(* IEC 61131-3 sources: STAR-PLC-Agent/results/raw/codex_matrix_resume_20261114/codex_deepseek/SELF007/functional/attempt_0001, 1 file *)

(* ---- test_program.st ---- *)
PROGRAM PLC_PRG
VAR
 BenchStep : UDINT := 0;
 BenchCalls : UDINT := 0;
 BenchDone : BOOL := FALSE;
 BenchUut0 : FB_Task;
 BenchUut1 : FB_Task;
 BenchUut2 : FB_Task;
 BenchUut3 : FB_Task;
 BenchUut4 : FB_Task;
 BenchUut5 : FB_Task;
 BenchUut6 : FB_Task;
 BenchUut7 : FB_Task;
 BenchUut8 : FB_Task;
 TraceIn_Demand : ARRAY[0..59] OF BOOL;
 TraceIn_FaultA : ARRAY[0..59] OF BOOL;
 TraceIn_FaultB : ARRAY[0..59] OF BOOL;
 TraceOut_PumpA : ARRAY[0..59] OF BOOL;
 TraceOut_PumpB : ARRAY[0..59] OF BOOL;
 TraceOut_LeadA : ARRAY[0..59] OF BOOL;
END_VAR

IF NOT BenchDone THEN
 CASE BenchStep OF
 0:
   BenchUut0.Demand := FALSE;
   BenchUut0.FaultA := FALSE;
   BenchUut0.FaultB := FALSE;
   TraceIn_Demand[0] := BenchUut0.Demand;
   TraceIn_FaultA[0] := BenchUut0.FaultA;
   TraceIn_FaultB[0] := BenchUut0.FaultB;
   BenchUut0();
   TraceOut_PumpA[0] := BenchUut0.PumpA;
   TraceOut_PumpB[0] := BenchUut0.PumpB;
   TraceOut_LeadA[0] := BenchUut0.LeadA;
   BenchCalls := BenchCalls + 1;
 1:
   BenchUut0.Demand := TRUE;
   BenchUut0.FaultA := FALSE;
   BenchUut0.FaultB := FALSE;
   TraceIn_Demand[1] := BenchUut0.Demand;
   TraceIn_FaultA[1] := BenchUut0.FaultA;
   TraceIn_FaultB[1] := BenchUut0.FaultB;
   BenchUut0();
   TraceOut_PumpA[1] := BenchUut0.PumpA;
   TraceOut_PumpB[1] := BenchUut0.PumpB;
   TraceOut_LeadA[1] := BenchUut0.LeadA;
   BenchCalls := BenchCalls + 1;
 2:
   BenchUut0.Demand := TRUE;
   BenchUut0.FaultA := FALSE;
   BenchUut0.FaultB := FALSE;
   TraceIn_Demand[2] := BenchUut0.Demand;
   TraceIn_FaultA[2] := BenchUut0.FaultA;
   TraceIn_FaultB[2] := BenchUut0.FaultB;
   BenchUut0();
   TraceOut_PumpA[2] := BenchUut0.PumpA;
   TraceOut_PumpB[2] := BenchUut0.PumpB;
   TraceOut_LeadA[2] := BenchUut0.LeadA;
   BenchCalls := BenchCalls + 1;
 3:
   BenchUut0.Demand := FALSE;
   BenchUut0.FaultA := FALSE;
   BenchUut0.FaultB := FALSE;
   TraceIn_Demand[3] := BenchUut0.Demand;
   TraceIn_FaultA[3] := BenchUut0.FaultA;
   TraceIn_FaultB[3] := BenchUut0.FaultB;
   BenchUut0();
   TraceOut_PumpA[3] := BenchUut0.PumpA;
   TraceOut_PumpB[3] := BenchUut0.PumpB;
   TraceOut_LeadA[3] := BenchUut0.LeadA;
   BenchCalls := BenchCalls + 1;
 4:
   BenchUut0.Demand := FALSE;
   BenchUut0.FaultA := FALSE;
   BenchUut0.FaultB := FALSE;
   TraceIn_Demand[4] := BenchUut0.Demand;
   TraceIn_FaultA[4] := BenchUut0.FaultA;
   TraceIn_FaultB[4] := BenchUut0.FaultB;
   BenchUut0();
   TraceOut_PumpA[4] := BenchUut0.PumpA;
   TraceOut_PumpB[4] := BenchUut0.PumpB;
   TraceOut_LeadA[4] := BenchUut0.LeadA;
   BenchCalls := BenchCalls + 1;
 5:
   BenchUut0.Demand := TRUE;
   BenchUut0.FaultA := FALSE;
   BenchUut0.FaultB := FALSE;
   TraceIn_Demand[5] := BenchUut0.Demand;
   TraceIn_FaultA[5] := BenchUut0.FaultA;
   TraceIn_FaultB[5] := BenchUut0.FaultB;
   BenchUut0();
   TraceOut_PumpA[5] := BenchUut0.PumpA;
   TraceOut_PumpB[5] := BenchUut0.PumpB;
   TraceOut_LeadA[5] := BenchUut0.LeadA;
   BenchCalls := BenchCalls + 1;
 6:
   BenchUut0.Demand := FALSE;
   BenchUut0.FaultA := FALSE;
   BenchUut0.FaultB := FALSE;
   TraceIn_Demand[6] := BenchUut0.Demand;
   TraceIn_FaultA[6] := BenchUut0.FaultA;
   TraceIn_FaultB[6] := BenchUut0.FaultB;
   BenchUut0();
   TraceOut_PumpA[6] := BenchUut0.PumpA;
   TraceOut_PumpB[6] := BenchUut0.PumpB;
   TraceOut_LeadA[6] := BenchUut0.LeadA;
   BenchCalls := BenchCalls + 1;
 7:
   BenchUut1.Demand := TRUE;
   BenchUut1.FaultA := TRUE;
   BenchUut1.FaultB := TRUE;
   TraceIn_Demand[7] := BenchUut1.Demand;
   TraceIn_FaultA[7] := BenchUut1.FaultA;
   TraceIn_FaultB[7] := BenchUut1.FaultB;
   BenchUut1();
   TraceOut_PumpA[7] := BenchUut1.PumpA;
   TraceOut_PumpB[7] := BenchUut1.PumpB;
   TraceOut_LeadA[7] := BenchUut1.LeadA;
   BenchCalls := BenchCalls + 1;
 8:
   BenchUut1.Demand := FALSE;
   BenchUut1.FaultA := TRUE;
   BenchUut1.FaultB := TRUE;
   TraceIn_Demand[8] := BenchUut1.Demand;
   TraceIn_FaultA[8] := BenchUut1.FaultA;
   TraceIn_FaultB[8] := BenchUut1.FaultB;
   BenchUut1();
   TraceOut_PumpA[8] := BenchUut1.PumpA;
   TraceOut_PumpB[8] := BenchUut1.PumpB;
   TraceOut_LeadA[8] := BenchUut1.LeadA;
   BenchCalls := BenchCalls + 1;
 9:
   BenchUut1.Demand := TRUE;
   BenchUut1.FaultA := TRUE;
   BenchUut1.FaultB := FALSE;
   TraceIn_Demand[9] := BenchUut1.Demand;
   TraceIn_FaultA[9] := BenchUut1.FaultA;
   TraceIn_FaultB[9] := BenchUut1.FaultB;
   BenchUut1();
   TraceOut_PumpA[9] := BenchUut1.PumpA;
   TraceOut_PumpB[9] := BenchUut1.PumpB;
   TraceOut_LeadA[9] := BenchUut1.LeadA;
   BenchCalls := BenchCalls + 1;
 10:
   BenchUut1.Demand := TRUE;
   BenchUut1.FaultA := FALSE;
   BenchUut1.FaultB := FALSE;
   TraceIn_Demand[10] := BenchUut1.Demand;
   TraceIn_FaultA[10] := BenchUut1.FaultA;
   TraceIn_FaultB[10] := BenchUut1.FaultB;
   BenchUut1();
   TraceOut_PumpA[10] := BenchUut1.PumpA;
   TraceOut_PumpB[10] := BenchUut1.PumpB;
   TraceOut_LeadA[10] := BenchUut1.LeadA;
   BenchCalls := BenchCalls + 1;
 11:
   BenchUut1.Demand := FALSE;
   BenchUut1.FaultA := TRUE;
   BenchUut1.FaultB := TRUE;
   TraceIn_Demand[11] := BenchUut1.Demand;
   TraceIn_FaultA[11] := BenchUut1.FaultA;
   TraceIn_FaultB[11] := BenchUut1.FaultB;
   BenchUut1();
   TraceOut_PumpA[11] := BenchUut1.PumpA;
   TraceOut_PumpB[11] := BenchUut1.PumpB;
   TraceOut_LeadA[11] := BenchUut1.LeadA;
   BenchCalls := BenchCalls + 1;
 12:
   BenchUut2.Demand := TRUE;
   BenchUut2.FaultA := TRUE;
   BenchUut2.FaultB := FALSE;
   TraceIn_Demand[12] := BenchUut2.Demand;
   TraceIn_FaultA[12] := BenchUut2.FaultA;
   TraceIn_FaultB[12] := BenchUut2.FaultB;
   BenchUut2();
   TraceOut_PumpA[12] := BenchUut2.PumpA;
   TraceOut_PumpB[12] := BenchUut2.PumpB;
   TraceOut_LeadA[12] := BenchUut2.LeadA;
   BenchCalls := BenchCalls + 1;
 13:
   BenchUut2.Demand := TRUE;
   BenchUut2.FaultA := TRUE;
   BenchUut2.FaultB := FALSE;
   TraceIn_Demand[13] := BenchUut2.Demand;
   TraceIn_FaultA[13] := BenchUut2.FaultA;
   TraceIn_FaultB[13] := BenchUut2.FaultB;
   BenchUut2();
   TraceOut_PumpA[13] := BenchUut2.PumpA;
   TraceOut_PumpB[13] := BenchUut2.PumpB;
   TraceOut_LeadA[13] := BenchUut2.LeadA;
   BenchCalls := BenchCalls + 1;
 14:
   BenchUut2.Demand := TRUE;
   BenchUut2.FaultA := TRUE;
   BenchUut2.FaultB := FALSE;
   TraceIn_Demand[14] := BenchUut2.Demand;
   TraceIn_FaultA[14] := BenchUut2.FaultA;
   TraceIn_FaultB[14] := BenchUut2.FaultB;
   BenchUut2();
   TraceOut_PumpA[14] := BenchUut2.PumpA;
   TraceOut_PumpB[14] := BenchUut2.PumpB;
   TraceOut_LeadA[14] := BenchUut2.LeadA;
   BenchCalls := BenchCalls + 1;
 15:
   BenchUut3.Demand := TRUE;
   BenchUut3.FaultA := FALSE;
   BenchUut3.FaultB := FALSE;
   TraceIn_Demand[15] := BenchUut3.Demand;
   TraceIn_FaultA[15] := BenchUut3.FaultA;
   TraceIn_FaultB[15] := BenchUut3.FaultB;
   BenchUut3();
   TraceOut_PumpA[15] := BenchUut3.PumpA;
   TraceOut_PumpB[15] := BenchUut3.PumpB;
   TraceOut_LeadA[15] := BenchUut3.LeadA;
   BenchCalls := BenchCalls + 1;
 16:
   BenchUut3.Demand := FALSE;
   BenchUut3.FaultA := FALSE;
   BenchUut3.FaultB := FALSE;
   TraceIn_Demand[16] := BenchUut3.Demand;
   TraceIn_FaultA[16] := BenchUut3.FaultA;
   TraceIn_FaultB[16] := BenchUut3.FaultB;
   BenchUut3();
   TraceOut_PumpA[16] := BenchUut3.PumpA;
   TraceOut_PumpB[16] := BenchUut3.PumpB;
   TraceOut_LeadA[16] := BenchUut3.LeadA;
   BenchCalls := BenchCalls + 1;
 17:
   BenchUut3.Demand := TRUE;
   BenchUut3.FaultA := FALSE;
   BenchUut3.FaultB := TRUE;
   TraceIn_Demand[17] := BenchUut3.Demand;
   TraceIn_FaultA[17] := BenchUut3.FaultA;
   TraceIn_FaultB[17] := BenchUut3.FaultB;
   BenchUut3();
   TraceOut_PumpA[17] := BenchUut3.PumpA;
   TraceOut_PumpB[17] := BenchUut3.PumpB;
   TraceOut_LeadA[17] := BenchUut3.LeadA;
   BenchCalls := BenchCalls + 1;
 18:
   BenchUut3.Demand := TRUE;
   BenchUut3.FaultA := TRUE;
   BenchUut3.FaultB := TRUE;
   TraceIn_Demand[18] := BenchUut3.Demand;
   TraceIn_FaultA[18] := BenchUut3.FaultA;
   TraceIn_FaultB[18] := BenchUut3.FaultB;
   BenchUut3();
   TraceOut_PumpA[18] := BenchUut3.PumpA;
   TraceOut_PumpB[18] := BenchUut3.PumpB;
   TraceOut_LeadA[18] := BenchUut3.LeadA;
   BenchCalls := BenchCalls + 1;
 19:
   BenchUut3.Demand := FALSE;
   BenchUut3.FaultA := TRUE;
   BenchUut3.FaultB := TRUE;
   TraceIn_Demand[19] := BenchUut3.Demand;
   TraceIn_FaultA[19] := BenchUut3.FaultA;
   TraceIn_FaultB[19] := BenchUut3.FaultB;
   BenchUut3();
   TraceOut_PumpA[19] := BenchUut3.PumpA;
   TraceOut_PumpB[19] := BenchUut3.PumpB;
   TraceOut_LeadA[19] := BenchUut3.LeadA;
   BenchCalls := BenchCalls + 1;
 20:
   BenchUut3.Demand := TRUE;
   BenchUut3.FaultA := FALSE;
   BenchUut3.FaultB := FALSE;
   TraceIn_Demand[20] := BenchUut3.Demand;
   TraceIn_FaultA[20] := BenchUut3.FaultA;
   TraceIn_FaultB[20] := BenchUut3.FaultB;
   BenchUut3();
   TraceOut_PumpA[20] := BenchUut3.PumpA;
   TraceOut_PumpB[20] := BenchUut3.PumpB;
   TraceOut_LeadA[20] := BenchUut3.LeadA;
   BenchCalls := BenchCalls + 1;
 21:
   BenchUut4.Demand := TRUE;
   BenchUut4.FaultA := FALSE;
   BenchUut4.FaultB := FALSE;
   TraceIn_Demand[21] := BenchUut4.Demand;
   TraceIn_FaultA[21] := BenchUut4.FaultA;
   TraceIn_FaultB[21] := BenchUut4.FaultB;
   BenchUut4();
   TraceOut_PumpA[21] := BenchUut4.PumpA;
   TraceOut_PumpB[21] := BenchUut4.PumpB;
   TraceOut_LeadA[21] := BenchUut4.LeadA;
   BenchCalls := BenchCalls + 1;
 22:
   BenchUut4.Demand := TRUE;
   BenchUut4.FaultA := TRUE;
   BenchUut4.FaultB := TRUE;
   TraceIn_Demand[22] := BenchUut4.Demand;
   TraceIn_FaultA[22] := BenchUut4.FaultA;
   TraceIn_FaultB[22] := BenchUut4.FaultB;
   BenchUut4();
   TraceOut_PumpA[22] := BenchUut4.PumpA;
   TraceOut_PumpB[22] := BenchUut4.PumpB;
   TraceOut_LeadA[22] := BenchUut4.LeadA;
   BenchCalls := BenchCalls + 1;
 23:
   BenchUut4.Demand := FALSE;
   BenchUut4.FaultA := TRUE;
   BenchUut4.FaultB := TRUE;
   TraceIn_Demand[23] := BenchUut4.Demand;
   TraceIn_FaultA[23] := BenchUut4.FaultA;
   TraceIn_FaultB[23] := BenchUut4.FaultB;
   BenchUut4();
   TraceOut_PumpA[23] := BenchUut4.PumpA;
   TraceOut_PumpB[23] := BenchUut4.PumpB;
   TraceOut_LeadA[23] := BenchUut4.LeadA;
   BenchCalls := BenchCalls + 1;
 24:
   BenchUut5.Demand := TRUE;
   BenchUut5.FaultA := FALSE;
   BenchUut5.FaultB := FALSE;
   TraceIn_Demand[24] := BenchUut5.Demand;
   TraceIn_FaultA[24] := BenchUut5.FaultA;
   TraceIn_FaultB[24] := BenchUut5.FaultB;
   BenchUut5();
   TraceOut_PumpA[24] := BenchUut5.PumpA;
   TraceOut_PumpB[24] := BenchUut5.PumpB;
   TraceOut_LeadA[24] := BenchUut5.LeadA;
   BenchCalls := BenchCalls + 1;
 25:
   BenchUut5.Demand := TRUE;
   BenchUut5.FaultA := TRUE;
   BenchUut5.FaultB := FALSE;
   TraceIn_Demand[25] := BenchUut5.Demand;
   TraceIn_FaultA[25] := BenchUut5.FaultA;
   TraceIn_FaultB[25] := BenchUut5.FaultB;
   BenchUut5();
   TraceOut_PumpA[25] := BenchUut5.PumpA;
   TraceOut_PumpB[25] := BenchUut5.PumpB;
   TraceOut_LeadA[25] := BenchUut5.LeadA;
   BenchCalls := BenchCalls + 1;
 26:
   BenchUut5.Demand := TRUE;
   BenchUut5.FaultA := FALSE;
   BenchUut5.FaultB := FALSE;
   TraceIn_Demand[26] := BenchUut5.Demand;
   TraceIn_FaultA[26] := BenchUut5.FaultA;
   TraceIn_FaultB[26] := BenchUut5.FaultB;
   BenchUut5();
   TraceOut_PumpA[26] := BenchUut5.PumpA;
   TraceOut_PumpB[26] := BenchUut5.PumpB;
   TraceOut_LeadA[26] := BenchUut5.LeadA;
   BenchCalls := BenchCalls + 1;
 27:
   BenchUut5.Demand := TRUE;
   BenchUut5.FaultA := TRUE;
   BenchUut5.FaultB := TRUE;
   TraceIn_Demand[27] := BenchUut5.Demand;
   TraceIn_FaultA[27] := BenchUut5.FaultA;
   TraceIn_FaultB[27] := BenchUut5.FaultB;
   BenchUut5();
   TraceOut_PumpA[27] := BenchUut5.PumpA;
   TraceOut_PumpB[27] := BenchUut5.PumpB;
   TraceOut_LeadA[27] := BenchUut5.LeadA;
   BenchCalls := BenchCalls + 1;
 28:
   BenchUut5.Demand := FALSE;
   BenchUut5.FaultA := TRUE;
   BenchUut5.FaultB := TRUE;
   TraceIn_Demand[28] := BenchUut5.Demand;
   TraceIn_FaultA[28] := BenchUut5.FaultA;
   TraceIn_FaultB[28] := BenchUut5.FaultB;
   BenchUut5();
   TraceOut_PumpA[28] := BenchUut5.PumpA;
   TraceOut_PumpB[28] := BenchUut5.PumpB;
   TraceOut_LeadA[28] := BenchUut5.LeadA;
   BenchCalls := BenchCalls + 1;
 29:
   BenchUut5.Demand := TRUE;
   BenchUut5.FaultA := FALSE;
   BenchUut5.FaultB := FALSE;
   TraceIn_Demand[29] := BenchUut5.Demand;
   TraceIn_FaultA[29] := BenchUut5.FaultA;
   TraceIn_FaultB[29] := BenchUut5.FaultB;
   BenchUut5();
   TraceOut_PumpA[29] := BenchUut5.PumpA;
   TraceOut_PumpB[29] := BenchUut5.PumpB;
   TraceOut_LeadA[29] := BenchUut5.LeadA;
   BenchCalls := BenchCalls + 1;
 30:
   BenchUut5.Demand := TRUE;
   BenchUut5.FaultA := FALSE;
   BenchUut5.FaultB := TRUE;
   TraceIn_Demand[30] := BenchUut5.Demand;
   TraceIn_FaultA[30] := BenchUut5.FaultA;
   TraceIn_FaultB[30] := BenchUut5.FaultB;
   BenchUut5();
   TraceOut_PumpA[30] := BenchUut5.PumpA;
   TraceOut_PumpB[30] := BenchUut5.PumpB;
   TraceOut_LeadA[30] := BenchUut5.LeadA;
   BenchCalls := BenchCalls + 1;
 31:
   BenchUut5.Demand := TRUE;
   BenchUut5.FaultA := FALSE;
   BenchUut5.FaultB := FALSE;
   TraceIn_Demand[31] := BenchUut5.Demand;
   TraceIn_FaultA[31] := BenchUut5.FaultA;
   TraceIn_FaultB[31] := BenchUut5.FaultB;
   BenchUut5();
   TraceOut_PumpA[31] := BenchUut5.PumpA;
   TraceOut_PumpB[31] := BenchUut5.PumpB;
   TraceOut_LeadA[31] := BenchUut5.LeadA;
   BenchCalls := BenchCalls + 1;
 32:
   BenchUut5.Demand := FALSE;
   BenchUut5.FaultA := FALSE;
   BenchUut5.FaultB := FALSE;
   TraceIn_Demand[32] := BenchUut5.Demand;
   TraceIn_FaultA[32] := BenchUut5.FaultA;
   TraceIn_FaultB[32] := BenchUut5.FaultB;
   BenchUut5();
   TraceOut_PumpA[32] := BenchUut5.PumpA;
   TraceOut_PumpB[32] := BenchUut5.PumpB;
   TraceOut_LeadA[32] := BenchUut5.LeadA;
   BenchCalls := BenchCalls + 1;
 33:
   BenchUut6.Demand := FALSE;
   BenchUut6.FaultA := FALSE;
   BenchUut6.FaultB := FALSE;
   TraceIn_Demand[33] := BenchUut6.Demand;
   TraceIn_FaultA[33] := BenchUut6.FaultA;
   TraceIn_FaultB[33] := BenchUut6.FaultB;
   BenchUut6();
   TraceOut_PumpA[33] := BenchUut6.PumpA;
   TraceOut_PumpB[33] := BenchUut6.PumpB;
   TraceOut_LeadA[33] := BenchUut6.LeadA;
   BenchCalls := BenchCalls + 1;
 34:
   BenchUut6.Demand := TRUE;
   BenchUut6.FaultA := FALSE;
   BenchUut6.FaultB := FALSE;
   TraceIn_Demand[34] := BenchUut6.Demand;
   TraceIn_FaultA[34] := BenchUut6.FaultA;
   TraceIn_FaultB[34] := BenchUut6.FaultB;
   BenchUut6();
   TraceOut_PumpA[34] := BenchUut6.PumpA;
   TraceOut_PumpB[34] := BenchUut6.PumpB;
   TraceOut_LeadA[34] := BenchUut6.LeadA;
   BenchCalls := BenchCalls + 1;
 35:
   BenchUut6.Demand := TRUE;
   BenchUut6.FaultA := FALSE;
   BenchUut6.FaultB := FALSE;
   TraceIn_Demand[35] := BenchUut6.Demand;
   TraceIn_FaultA[35] := BenchUut6.FaultA;
   TraceIn_FaultB[35] := BenchUut6.FaultB;
   BenchUut6();
   TraceOut_PumpA[35] := BenchUut6.PumpA;
   TraceOut_PumpB[35] := BenchUut6.PumpB;
   TraceOut_LeadA[35] := BenchUut6.LeadA;
   BenchCalls := BenchCalls + 1;
 36:
   BenchUut6.Demand := FALSE;
   BenchUut6.FaultA := FALSE;
   BenchUut6.FaultB := FALSE;
   TraceIn_Demand[36] := BenchUut6.Demand;
   TraceIn_FaultA[36] := BenchUut6.FaultA;
   TraceIn_FaultB[36] := BenchUut6.FaultB;
   BenchUut6();
   TraceOut_PumpA[36] := BenchUut6.PumpA;
   TraceOut_PumpB[36] := BenchUut6.PumpB;
   TraceOut_LeadA[36] := BenchUut6.LeadA;
   BenchCalls := BenchCalls + 1;
 37:
   BenchUut6.Demand := FALSE;
   BenchUut6.FaultA := FALSE;
   BenchUut6.FaultB := FALSE;
   TraceIn_Demand[37] := BenchUut6.Demand;
   TraceIn_FaultA[37] := BenchUut6.FaultA;
   TraceIn_FaultB[37] := BenchUut6.FaultB;
   BenchUut6();
   TraceOut_PumpA[37] := BenchUut6.PumpA;
   TraceOut_PumpB[37] := BenchUut6.PumpB;
   TraceOut_LeadA[37] := BenchUut6.LeadA;
   BenchCalls := BenchCalls + 1;
 38:
   BenchUut6.Demand := TRUE;
   BenchUut6.FaultA := FALSE;
   BenchUut6.FaultB := FALSE;
   TraceIn_Demand[38] := BenchUut6.Demand;
   TraceIn_FaultA[38] := BenchUut6.FaultA;
   TraceIn_FaultB[38] := BenchUut6.FaultB;
   BenchUut6();
   TraceOut_PumpA[38] := BenchUut6.PumpA;
   TraceOut_PumpB[38] := BenchUut6.PumpB;
   TraceOut_LeadA[38] := BenchUut6.LeadA;
   BenchCalls := BenchCalls + 1;
 39:
   BenchUut6.Demand := FALSE;
   BenchUut6.FaultA := FALSE;
   BenchUut6.FaultB := FALSE;
   TraceIn_Demand[39] := BenchUut6.Demand;
   TraceIn_FaultA[39] := BenchUut6.FaultA;
   TraceIn_FaultB[39] := BenchUut6.FaultB;
   BenchUut6();
   TraceOut_PumpA[39] := BenchUut6.PumpA;
   TraceOut_PumpB[39] := BenchUut6.PumpB;
   TraceOut_LeadA[39] := BenchUut6.LeadA;
   BenchCalls := BenchCalls + 1;
 40:
   BenchUut6.Demand := TRUE;
   BenchUut6.FaultA := FALSE;
   BenchUut6.FaultB := FALSE;
   TraceIn_Demand[40] := BenchUut6.Demand;
   TraceIn_FaultA[40] := BenchUut6.FaultA;
   TraceIn_FaultB[40] := BenchUut6.FaultB;
   BenchUut6();
   TraceOut_PumpA[40] := BenchUut6.PumpA;
   TraceOut_PumpB[40] := BenchUut6.PumpB;
   TraceOut_LeadA[40] := BenchUut6.LeadA;
   BenchCalls := BenchCalls + 1;
 41:
   BenchUut6.Demand := TRUE;
   BenchUut6.FaultA := FALSE;
   BenchUut6.FaultB := FALSE;
   TraceIn_Demand[41] := BenchUut6.Demand;
   TraceIn_FaultA[41] := BenchUut6.FaultA;
   TraceIn_FaultB[41] := BenchUut6.FaultB;
   BenchUut6();
   TraceOut_PumpA[41] := BenchUut6.PumpA;
   TraceOut_PumpB[41] := BenchUut6.PumpB;
   TraceOut_LeadA[41] := BenchUut6.LeadA;
   BenchCalls := BenchCalls + 1;
 42:
   BenchUut7.Demand := FALSE;
   BenchUut7.FaultA := FALSE;
   BenchUut7.FaultB := FALSE;
   TraceIn_Demand[42] := BenchUut7.Demand;
   TraceIn_FaultA[42] := BenchUut7.FaultA;
   TraceIn_FaultB[42] := BenchUut7.FaultB;
   BenchUut7();
   TraceOut_PumpA[42] := BenchUut7.PumpA;
   TraceOut_PumpB[42] := BenchUut7.PumpB;
   TraceOut_LeadA[42] := BenchUut7.LeadA;
   BenchCalls := BenchCalls + 1;
 43:
   BenchUut7.Demand := TRUE;
   BenchUut7.FaultA := FALSE;
   BenchUut7.FaultB := FALSE;
   TraceIn_Demand[43] := BenchUut7.Demand;
   TraceIn_FaultA[43] := BenchUut7.FaultA;
   TraceIn_FaultB[43] := BenchUut7.FaultB;
   BenchUut7();
   TraceOut_PumpA[43] := BenchUut7.PumpA;
   TraceOut_PumpB[43] := BenchUut7.PumpB;
   TraceOut_LeadA[43] := BenchUut7.LeadA;
   BenchCalls := BenchCalls + 1;
 44:
   BenchUut7.Demand := TRUE;
   BenchUut7.FaultA := FALSE;
   BenchUut7.FaultB := FALSE;
   TraceIn_Demand[44] := BenchUut7.Demand;
   TraceIn_FaultA[44] := BenchUut7.FaultA;
   TraceIn_FaultB[44] := BenchUut7.FaultB;
   BenchUut7();
   TraceOut_PumpA[44] := BenchUut7.PumpA;
   TraceOut_PumpB[44] := BenchUut7.PumpB;
   TraceOut_LeadA[44] := BenchUut7.LeadA;
   BenchCalls := BenchCalls + 1;
 45:
   BenchUut7.Demand := FALSE;
   BenchUut7.FaultA := FALSE;
   BenchUut7.FaultB := FALSE;
   TraceIn_Demand[45] := BenchUut7.Demand;
   TraceIn_FaultA[45] := BenchUut7.FaultA;
   TraceIn_FaultB[45] := BenchUut7.FaultB;
   BenchUut7();
   TraceOut_PumpA[45] := BenchUut7.PumpA;
   TraceOut_PumpB[45] := BenchUut7.PumpB;
   TraceOut_LeadA[45] := BenchUut7.LeadA;
   BenchCalls := BenchCalls + 1;
 46:
   BenchUut7.Demand := FALSE;
   BenchUut7.FaultA := FALSE;
   BenchUut7.FaultB := FALSE;
   TraceIn_Demand[46] := BenchUut7.Demand;
   TraceIn_FaultA[46] := BenchUut7.FaultA;
   TraceIn_FaultB[46] := BenchUut7.FaultB;
   BenchUut7();
   TraceOut_PumpA[46] := BenchUut7.PumpA;
   TraceOut_PumpB[46] := BenchUut7.PumpB;
   TraceOut_LeadA[46] := BenchUut7.LeadA;
   BenchCalls := BenchCalls + 1;
 47:
   BenchUut7.Demand := TRUE;
   BenchUut7.FaultA := FALSE;
   BenchUut7.FaultB := FALSE;
   TraceIn_Demand[47] := BenchUut7.Demand;
   TraceIn_FaultA[47] := BenchUut7.FaultA;
   TraceIn_FaultB[47] := BenchUut7.FaultB;
   BenchUut7();
   TraceOut_PumpA[47] := BenchUut7.PumpA;
   TraceOut_PumpB[47] := BenchUut7.PumpB;
   TraceOut_LeadA[47] := BenchUut7.LeadA;
   BenchCalls := BenchCalls + 1;
 48:
   BenchUut7.Demand := FALSE;
   BenchUut7.FaultA := FALSE;
   BenchUut7.FaultB := FALSE;
   TraceIn_Demand[48] := BenchUut7.Demand;
   TraceIn_FaultA[48] := BenchUut7.FaultA;
   TraceIn_FaultB[48] := BenchUut7.FaultB;
   BenchUut7();
   TraceOut_PumpA[48] := BenchUut7.PumpA;
   TraceOut_PumpB[48] := BenchUut7.PumpB;
   TraceOut_LeadA[48] := BenchUut7.LeadA;
   BenchCalls := BenchCalls + 1;
 49:
   BenchUut7.Demand := FALSE;
   BenchUut7.FaultA := TRUE;
   BenchUut7.FaultB := FALSE;
   TraceIn_Demand[49] := BenchUut7.Demand;
   TraceIn_FaultA[49] := BenchUut7.FaultA;
   TraceIn_FaultB[49] := BenchUut7.FaultB;
   BenchUut7();
   TraceOut_PumpA[49] := BenchUut7.PumpA;
   TraceOut_PumpB[49] := BenchUut7.PumpB;
   TraceOut_LeadA[49] := BenchUut7.LeadA;
   BenchCalls := BenchCalls + 1;
 50:
   BenchUut7.Demand := FALSE;
   BenchUut7.FaultA := TRUE;
   BenchUut7.FaultB := FALSE;
   TraceIn_Demand[50] := BenchUut7.Demand;
   TraceIn_FaultA[50] := BenchUut7.FaultA;
   TraceIn_FaultB[50] := BenchUut7.FaultB;
   BenchUut7();
   TraceOut_PumpA[50] := BenchUut7.PumpA;
   TraceOut_PumpB[50] := BenchUut7.PumpB;
   TraceOut_LeadA[50] := BenchUut7.LeadA;
   BenchCalls := BenchCalls + 1;
 51:
   BenchUut8.Demand := FALSE;
   BenchUut8.FaultA := FALSE;
   BenchUut8.FaultB := FALSE;
   TraceIn_Demand[51] := BenchUut8.Demand;
   TraceIn_FaultA[51] := BenchUut8.FaultA;
   TraceIn_FaultB[51] := BenchUut8.FaultB;
   BenchUut8();
   TraceOut_PumpA[51] := BenchUut8.PumpA;
   TraceOut_PumpB[51] := BenchUut8.PumpB;
   TraceOut_LeadA[51] := BenchUut8.LeadA;
   BenchCalls := BenchCalls + 1;
 52:
   BenchUut8.Demand := TRUE;
   BenchUut8.FaultA := FALSE;
   BenchUut8.FaultB := FALSE;
   TraceIn_Demand[52] := BenchUut8.Demand;
   TraceIn_FaultA[52] := BenchUut8.FaultA;
   TraceIn_FaultB[52] := BenchUut8.FaultB;
   BenchUut8();
   TraceOut_PumpA[52] := BenchUut8.PumpA;
   TraceOut_PumpB[52] := BenchUut8.PumpB;
   TraceOut_LeadA[52] := BenchUut8.LeadA;
   BenchCalls := BenchCalls + 1;
 53:
   BenchUut8.Demand := TRUE;
   BenchUut8.FaultA := FALSE;
   BenchUut8.FaultB := FALSE;
   TraceIn_Demand[53] := BenchUut8.Demand;
   TraceIn_FaultA[53] := BenchUut8.FaultA;
   TraceIn_FaultB[53] := BenchUut8.FaultB;
   BenchUut8();
   TraceOut_PumpA[53] := BenchUut8.PumpA;
   TraceOut_PumpB[53] := BenchUut8.PumpB;
   TraceOut_LeadA[53] := BenchUut8.LeadA;
   BenchCalls := BenchCalls + 1;
 54:
   BenchUut8.Demand := FALSE;
   BenchUut8.FaultA := FALSE;
   BenchUut8.FaultB := FALSE;
   TraceIn_Demand[54] := BenchUut8.Demand;
   TraceIn_FaultA[54] := BenchUut8.FaultA;
   TraceIn_FaultB[54] := BenchUut8.FaultB;
   BenchUut8();
   TraceOut_PumpA[54] := BenchUut8.PumpA;
   TraceOut_PumpB[54] := BenchUut8.PumpB;
   TraceOut_LeadA[54] := BenchUut8.LeadA;
   BenchCalls := BenchCalls + 1;
 55:
   BenchUut8.Demand := FALSE;
   BenchUut8.FaultA := FALSE;
   BenchUut8.FaultB := FALSE;
   TraceIn_Demand[55] := BenchUut8.Demand;
   TraceIn_FaultA[55] := BenchUut8.FaultA;
   TraceIn_FaultB[55] := BenchUut8.FaultB;
   BenchUut8();
   TraceOut_PumpA[55] := BenchUut8.PumpA;
   TraceOut_PumpB[55] := BenchUut8.PumpB;
   TraceOut_LeadA[55] := BenchUut8.LeadA;
   BenchCalls := BenchCalls + 1;
 56:
   BenchUut8.Demand := TRUE;
   BenchUut8.FaultA := FALSE;
   BenchUut8.FaultB := FALSE;
   TraceIn_Demand[56] := BenchUut8.Demand;
   TraceIn_FaultA[56] := BenchUut8.FaultA;
   TraceIn_FaultB[56] := BenchUut8.FaultB;
   BenchUut8();
   TraceOut_PumpA[56] := BenchUut8.PumpA;
   TraceOut_PumpB[56] := BenchUut8.PumpB;
   TraceOut_LeadA[56] := BenchUut8.LeadA;
   BenchCalls := BenchCalls + 1;
 57:
   BenchUut8.Demand := FALSE;
   BenchUut8.FaultA := FALSE;
   BenchUut8.FaultB := FALSE;
   TraceIn_Demand[57] := BenchUut8.Demand;
   TraceIn_FaultA[57] := BenchUut8.FaultA;
   TraceIn_FaultB[57] := BenchUut8.FaultB;
   BenchUut8();
   TraceOut_PumpA[57] := BenchUut8.PumpA;
   TraceOut_PumpB[57] := BenchUut8.PumpB;
   TraceOut_LeadA[57] := BenchUut8.LeadA;
   BenchCalls := BenchCalls + 1;
 58:
   BenchUut8.Demand := FALSE;
   BenchUut8.FaultA := FALSE;
   BenchUut8.FaultB := TRUE;
   TraceIn_Demand[58] := BenchUut8.Demand;
   TraceIn_FaultA[58] := BenchUut8.FaultA;
   TraceIn_FaultB[58] := BenchUut8.FaultB;
   BenchUut8();
   TraceOut_PumpA[58] := BenchUut8.PumpA;
   TraceOut_PumpB[58] := BenchUut8.PumpB;
   TraceOut_LeadA[58] := BenchUut8.LeadA;
   BenchCalls := BenchCalls + 1;
 59:
   BenchUut8.Demand := FALSE;
   BenchUut8.FaultA := FALSE;
   BenchUut8.FaultB := TRUE;
   TraceIn_Demand[59] := BenchUut8.Demand;
   TraceIn_FaultA[59] := BenchUut8.FaultA;
   TraceIn_FaultB[59] := BenchUut8.FaultB;
   BenchUut8();
   TraceOut_PumpA[59] := BenchUut8.PumpA;
   TraceOut_PumpB[59] := BenchUut8.PumpB;
   TraceOut_LeadA[59] := BenchUut8.LeadA;
   BenchCalls := BenchCalls + 1;
 END_CASE;
 BenchStep := BenchStep + 1;
 IF BenchStep >= 60 THEN BenchDone := TRUE; END_IF;
END_IF;
END_PROGRAM
